// TIA Portal V19 export
// export: Created 2026-10-16T08:35:17.5230422Z, ExportSetting WithDefaults, DisplayName Totally Integrated Automation Portal, DisplayVersion V19, DisplayName TIA Portal Openness, DisplayVersion V19, DisplayName TIA Portal Version Control Interface, DisplayVersion V19, DisplayName STEP 7 Professional, DisplayVersion V19, DisplayName STEP 7 Safety, DisplayVersion V19, DisplayName WinCC Basic/Comfort/Advanced, DisplayVersion V19, DisplayName WinCC Unified, DisplayVersion V19
Screen "WZOR_ROLL"  800x480, Number=1
  ScreenLayer 
    Button "Button_1" at 215,36 size 96x32  Mode=Text, TextOff="Test", TextOn="Text"
      on Press: SetBit(Tag := WzorPrzycisk)
      on Release: ResetBit(Tag := WzorPrzycisk)
    IOField "I/O field_1" at 345,36 size 96x32  DataFormat=Decimal, FormatPattern=s99999, Mode=InOutput
      ProcessValue := WzorLiczba
    TextField "Text field_1" at 118,48 size 84x20  Text="Wzór ROLL"
    Circle "Circle_1" at 584,36 size 48x48
      RangeAppearanceAnimation "RangeAppearanceAnimation"
        tag WzorStan
        0..0: back #d9d9d9, fore #181c31
        1..1: back #339966, fore #181c31
